# EPICS substitutions: db/Beckhoff_7XXX/ecmcEX72XX_OPT_encoderStatus.substitutions
file "ecmcEL72XX_FB_STAT.template"
{
  pattern {CH_ID}
          {"$(OPT_CH_ID=01)"}
}
